Yaskawa INFORM job: 20211127CHUKOUOFFLINE.JBI

/JOB
//NAME 20211127CHUKOUOFFLINE
//POS
///NPOS 6,0,6,0,0,0
///TOOL 1
///POSTYPE PULSE
///PULSE
C00000=-4685,43412,27733,-3116,-80596,2914
C00001=-4299,32992,-15629,-4269,-52439,3794
C00002=-4299,32992,-15629,-4269,-52439,3794
C00003=-4299,32992,-15629,-4269,-52439,3794
C00004=-4299,32992,-15629,-4269,-52439,3794
C00005=-4079,36005,21062,-3522,-75393,2906
///TOOL 0
EC00000=-4,-74112
EC00001=-4,-74112
EC00002=-4,-74112
EC00003=-4,-169112
EC00004=-4,-313392
EC00005=-4,-313392
//INST
///DATE 2021/11/27 18:52
///ATTR SC,RW
///GROUP1 RB1
///GROUP2 ST1
NOP
MOVJ C00000 VJ=10.00  +MOVJ EC00000 VJ=10.00
MOVL C00001 V=20.0  +MOVJ EC00001 VJ=10.00
CALL JOB:SAVETRAJ
SMOVC C00002 V=5.0  +MOVJ EC00002
SMOVC C00003 V=5.0  +MOVJ EC00003
SMOVC C00004 V=5.0  +MOVJ EC00004
CALL JOB:ENDTRAJ
MOVL C00005 V=20.0  +MOVJ EC00005 VJ=10.00
END
